(* PLC project webui_demo, Tether tplc *)

PROGRAM MAIN
  VAR_INPUT
    Limit : ? := 90;
  END_VAR
  VAR
    Start AT %IX0.0 : ?;
    Heat AT %QX0.0 : ?;
  END_VAR
  VAR
    T1 : ?;
  END_VAR

(* FBD diagram, written out as Structured Text *)
END_PROGRAM
